Staubli VAL3: exercice2.pgx

program exercice2()
begin
  movej(jDepart,tPince,mRapide)
  call ouvrirPince()
  movej(appro(Prise5[0],{0,0,-50,0,0,0}),tPince,mRapide)
  movel(Prise5[0],tPince,mLent)
  call fermerPince()
  movel(appro(Prise5[0],{0,0,-50,0,0,0}),tPince,mRapide)

  movej(jDepart,tPince,mRapide)
  movej(appro(pDepose[0],{0,0,-50,0,0,0}),tPince,mRapide)
  movel(pDepose[0],tPince,mLent)
  call ouvrirPince()
  movel(appro(pDepose,{0,0,-50,0,0,0}),tPince,mRapide)

  movej(jDepart,tPince,mLent)

  waitEndMove()
end
